// TIA Portal V21 export
// export: Created 2000-01-01T00:00:00.0000000Z, ExportSetting None
TYPE "UDT_HMI_FIO_Turntable"
   STRUCT
      bManualMode { ExternalWritable := 'False'} : Bool;   // TRUE手动, FALSE自动
      bStartCmd { ExternalWritable := 'False'} : Bool;   // HMI启动命令
      bStopCmd { ExternalWritable := 'False'} : Bool;   // HMI停止命令
      bResetCmd { ExternalWritable := 'False'} : Bool;   // HMI故障复位
      bRouteTo90Deg { ExternalWritable := 'False'} : Bool;   // 分流路由选择：TRUE=旋转90度侧向出料, FALSE=0度直通出料
      bManualTurn { ExternalWritable := 'False'} : Bool;   // 手动驱动转盘旋转至90度
      bManualRollPlus { ExternalWritable := 'False'} : Bool;   // 手动驱动转盘滚筒正转
      tActionTimeout { ExternalWritable := 'False'} : Time;   // 转盘旋转/进出料超时时间（默认 T#5s）
      iCurrentStep { ExternalWritable := 'False'} : Int;   // 状态反馈：当前步序
      diRoutedCount { ExternalWritable := 'False'} : DInt;   // 状态反馈：累计通过托盘数
      bFault { ExternalWritable := 'False'} : Bool;   // 状态反馈：故障标志
      wStatus { ExternalWritable := 'False'} : Word;   // 状态码：16#0000正常, 16#7000待机, 16#8401转盘动作超时, 16#8402急停触发
   END_STRUCT;
END_TYPE
